Fanuc KAREL source: KO00037.KL

PROGRAM KO00037
%NOLOCKGROUP
%ENVIRONMENT MIR
VAR
  P1: POSITION
  P2: XYZWPR
  F: BOOLEAN
  OUT: POSITION
BEGIN
  F = TRUE
  OUT = MIRROR(P1, P2, F)
END KO00037
